// TIA Portal V20 export
TYPE "Wartungszähler_Zyklen"
   STRUCT
      Gesamtzyklen : DInt;
      Zyklen_soll : DInt;
      Zyklen_seit_Wartung : DInt;
      Zyklen_bis_Wartung : DInt;
      Zähler_reset : Bool;
      SM_Wartung_fällig : Bool;
   END_STRUCT;
END_TYPE
